Fanuc KAREL source: kt00024.KL

-- PROVISIONAL review KL for V770-1; original PC SHA256 ad4d2fa41dc6ec79eabcdff8a8b8ceb0e47e22b11b8e4214befd5fcf75bc7cc8
-- Incomplete behavior may be omitted. Consult companion uncertainty JSON. Do not deploy.
PROGRAM KT00024
%NOLOCKGROUP
VAR
  OUT : REAL
-- UNRESOLVED_DECL Y1 type=002018
-- UNRESOLVED_DECL H2 type=002017
BEGIN
  -- UNRESOLVED_PC offsets 5-19; opcodes 2E,22,9D,33,B2
  -- UNRESOLVED_PC offsets 24-38; opcodes 2E,22,9D,33,B4
  -- UNRESOLVED_PC offsets 43-69; opcodes 22,9D,33,B1,22,9D,33,B3,52,64,23
  -- UNRESOLVED_PC offsets 74-78; opcodes 7F
END KT00024
